FUNCTION_BLOCK FB_StrokeStation
VAR_OUTPUT
    Phase : DINT; // Outstroke 0..100, return 101..200
    Done : BOOL;
END_VAR
VAR
    Cylinder : FB_VirtualCylinder;
    Returning : BOOL;
END_VAR

METHOD ResetStation
Cylinder.Home();
Returning := FALSE;
Phase := 0;
Done := FALSE;
END_METHOD

METHOD Step
IF Done THEN RETURN; END_IF
Cylinder.FollowStroke(Forward := NOT Returning);
IF Returning THEN
    Phase := 200 - Cylinder.Position;
    Done := Cylinder.Position = 0;
ELSE
    Phase := Cylinder.Position;
    Returning := Cylinder.Position = 100;
END_IF
END_METHOD

END_FUNCTION_BLOCK

(* stored: Version 1.1.0.1, ProductVersion 3.1.4024.53
   POU FB_StrokeStation: Id {52592E20-A431-4FDA-93CC-000000000010}
   Method ResetStation: Id {52592E20-A431-4FDA-93CC-000000000008}
   Method Step: Id {52592E20-A431-4FDA-93CC-000000000009} *)
